(* IEC 61131-3 sources: rsb-lab/vlan50/plc-programs, 6 files *)

(* ---- brewhouse.st ---- *)
PROGRAM plc_prg
VAR
    MashTemp           AT %QW0 : INT;
    MashLevel          AT %QW1 : INT;
    MashPH             AT %QW2 : INT;
    LauterTurbidity    AT %QW3 : INT;
    LauterLevel        AT %QW4 : INT;
    KettleTemp         AT %QW5 : INT;
    KettleLevel        AT %QW6 : INT;
    KettlePressure     AT %QW7 : INT;
    WhirlpoolTemp      AT %QW8 : INT;
    ChillerOutTemp     AT %QW9 : INT;

    MashAgitator       AT %QX0.0 : BOOL;
    MashOutlet         AT %QX0.1 : BOOL;
    LauterToKettle     AT %QX0.2 : BOOL;
    LauterRecirculate  AT %QX0.3 : BOOL;
    KettleSteam        AT %QX0.4 : BOOL;
    KettleToWhirlpool  AT %QX0.5 : BOOL;
    WhirlpoolOutlet    AT %QX0.6 : BOOL;
    ChillerOutlet      AT %QX0.7 : BOOL;

    AlarmTurbidity     AT %QX1.0 : BOOL;  (* coil 8 *)
    AlarmKettleTemp    AT %QX1.1 : BOOL;  (* coil 9 *)
    AlarmKettlePress   AT %QX1.2 : BOOL;  (* coil 10 *)
    AlarmChillerTemp   AT %QX1.3 : BOOL;  (* coil 11 *)
    WhirlpoolReady     AT %QX1.4 : BOOL;  (* coil 12 *)
END_VAR
VAR
    TransferSeen : BOOL;
    WhirlpoolRest : TON;
END_VAR

AlarmTurbidity   := LauterTurbidity > 200;
AlarmKettleTemp  := KettleTemp >= 1000;
AlarmKettlePress := KettlePressure >= 1200;
AlarmChillerTemp := ChillerOutTemp > 200;

IF AlarmTurbidity AND (LauterLevel > 2) THEN
    LauterToKettle := FALSE;
    LauterRecirculate := TRUE;
ELSIF LauterLevel <= 2 THEN
    LauterToKettle := FALSE;
    LauterRecirculate := FALSE;
END_IF;

IF AlarmKettleTemp OR AlarmKettlePress THEN
    KettleSteam := FALSE;
END_IF;

IF KettleToWhirlpool THEN
    TransferSeen := TRUE;
END_IF;

WhirlpoolRest(IN := TransferSeen AND NOT KettleToWhirlpool, PT := T#20m);
WhirlpoolReady := WhirlpoolRest.Q;

IF NOT WhirlpoolReady THEN
    WhirlpoolOutlet := FALSE;
END_IF;

IF AlarmChillerTemp THEN
    ChillerOutlet := FALSE;
END_IF;

IF ChillerOutlet AND (ChillerOutTemp <= 200) THEN
    TransferSeen := FALSE;
END_IF;

END_PROGRAM

CONFIGURATION Config0
    RESOURCE Res0 ON PLC
        TASK task0(INTERVAL := T#100ms, PRIORITY := 0);
        PROGRAM instance0 WITH task0 : plc_prg;
    END_RESOURCE
END_CONFIGURATION

(* ---- conditioning.st ---- *)
PROGRAM plc_prg
VAR
    BBT1Temp       AT %QW0 : INT;
    BBT1Pressure   AT %QW1 : INT;
    BBT1Level      AT %QW2 : INT;
    BBT1Turbidity  AT %QW3 : INT;
    BBT2Temp       AT %QW10 : INT;
    BBT2Pressure   AT %QW11 : INT;
    BBT2Level      AT %QW12 : INT;
    BBT2Turbidity  AT %QW13 : INT;

    BBT1Glycol     AT %QX0.0 : BOOL;
    BBT1CO2Dose    AT %QX0.1 : BOOL;
    BBT1Outlet     AT %QX0.2 : BOOL;
    BBT1Vent       AT %QX0.3 : BOOL;
    BBT2Glycol     AT %QX1.2 : BOOL;
    BBT2CO2Dose    AT %QX1.3 : BOOL;
    BBT2Outlet     AT %QX1.4 : BOOL;
    BBT2Vent       AT %QX1.5 : BOOL;

    AlarmBBT1Temp      AT %QX2.4 : BOOL; (* coil 20 *)
    AlarmBBT2Temp      AT %QX2.5 : BOOL; (* coil 21 *)
    AlarmBBT1Pressure  AT %QX2.6 : BOOL; (* coil 22 *)
    AlarmBBT2Pressure  AT %QX2.7 : BOOL; (* coil 23 *)
    BBT1Ready          AT %QX3.0 : BOOL; (* coil 24 *)
    BBT2Ready          AT %QX3.1 : BOOL; (* coil 25 *)
END_VAR
VAR
    BBT1StableTimer : TON;
    BBT2StableTimer : TON;
END_VAR

AlarmBBT1Temp := BBT1Temp > 20;
AlarmBBT2Temp := BBT2Temp > 20;
AlarmBBT1Pressure := BBT1Pressure > 2000;
AlarmBBT2Pressure := BBT2Pressure > 2000;

IF BBT1Temp > 20 THEN BBT1Glycol := TRUE; ELSIF BBT1Temp <= 0 THEN BBT1Glycol := FALSE; END_IF;
IF BBT2Temp > 20 THEN BBT2Glycol := TRUE; ELSIF BBT2Temp <= 0 THEN BBT2Glycol := FALSE; END_IF;

IF BBT1Pressure > 2000 THEN BBT1CO2Dose := FALSE; END_IF;
IF BBT2Pressure > 2000 THEN BBT2CO2Dose := FALSE; END_IF;

IF BBT1Pressure >= 2500 THEN BBT1Vent := TRUE; ELSIF BBT1Pressure < 2200 THEN BBT1Vent := FALSE; END_IF;
IF BBT2Pressure >= 2500 THEN BBT2Vent := TRUE; ELSIF BBT2Pressure < 2200 THEN BBT2Vent := FALSE; END_IF;

BBT1StableTimer(IN := (BBT1Temp >= 0) AND (BBT1Temp <= 20) AND (BBT1Turbidity <= 20), PT := T#10m);
BBT2StableTimer(IN := (BBT2Temp >= 0) AND (BBT2Temp <= 20) AND (BBT2Turbidity <= 20), PT := T#10m);
BBT1Ready := BBT1StableTimer.Q;
BBT2Ready := BBT2StableTimer.Q;

IF NOT BBT1Ready THEN BBT1Outlet := FALSE; END_IF;
IF NOT BBT2Ready THEN BBT2Outlet := FALSE; END_IF;

IF BBT1Level <= 2 THEN BBT1Outlet := FALSE; END_IF;
IF BBT2Level <= 2 THEN BBT2Outlet := FALSE; END_IF;

END_PROGRAM

CONFIGURATION Config0
    RESOURCE Res0 ON PLC
        TASK task0(INTERVAL := T#100ms, PRIORITY := 0);
        PROGRAM instance0 WITH task0 : plc_prg;
    END_RESOURCE
END_CONFIGURATION

(* ---- fermentation.st ---- *)
PROGRAM plc_prg
VAR
    T1Temp       AT %QW0 : INT;
    T1Pressure   AT %QW1 : INT;
    T1Level      AT %QW2 : INT;
    T1PH         AT %QW3 : INT;
    CO2Header    AT %QW4 : INT;
    CO2Flow      AT %QW5 : INT;

    T2Temp       AT %QW10 : INT;
    T2Pressure   AT %QW11 : INT;
    T2Level      AT %QW12 : INT;
    T2PH         AT %QW13 : INT;
    T3Temp       AT %QW20 : INT;
    T3Pressure   AT %QW21 : INT;
    T3Level      AT %QW22 : INT;
    T3PH         AT %QW23 : INT;
    T4Temp       AT %QW30 : INT;
    T4Pressure   AT %QW31 : INT;
    T4Level      AT %QW32 : INT;
    T4PH         AT %QW33 : INT;

    T1Glycol     AT %QX0.0 : BOOL;
    T1Outlet     AT %QX0.1 : BOOL;
    T1CIP        AT %QX0.2 : BOOL;
    T2Glycol     AT %QX1.2 : BOOL;
    T2Outlet     AT %QX1.3 : BOOL;
    T2CIP        AT %QX1.4 : BOOL;
    T3Glycol     AT %QX2.4 : BOOL;
    T3Outlet     AT %QX2.5 : BOOL;
    T3CIP        AT %QX2.6 : BOOL;
    T4Glycol     AT %QX3.6 : BOOL;
    T4Outlet     AT %QX3.7 : BOOL;
    T4CIP        AT %QX4.0 : BOOL;
    CO2Vent      AT %QX5.0 : BOOL;
    CO2Recovery  AT %QX5.1 : BOOL;

    AlarmHighPressure AT %QX6.2 : BOOL; (* coil 50 *)
    AlarmEmergency    AT %QX6.3 : BOOL; (* coil 51 *)
    T1Complete        AT %QX6.4 : BOOL; (* coil 52 *)
    T2Complete        AT %QX6.5 : BOOL; (* coil 53 *)
    T3Complete        AT %QX6.6 : BOOL; (* coil 54 *)
    T4Complete        AT %QX6.7 : BOOL; (* coil 55 *)
END_VAR
VAR
    T1FermentTimer : TON;
    T2FermentTimer : TON;
    T3FermentTimer : TON;
    T4FermentTimer : TON;
END_VAR

IF T1Temp > 205 THEN T1Glycol := TRUE; ELSIF T1Temp < 195 THEN T1Glycol := FALSE; END_IF;
IF T2Temp > 205 THEN T2Glycol := TRUE; ELSIF T2Temp < 195 THEN T2Glycol := FALSE; END_IF;
IF T3Temp > 205 THEN T3Glycol := TRUE; ELSIF T3Temp < 195 THEN T3Glycol := FALSE; END_IF;
IF T4Temp > 205 THEN T4Glycol := TRUE; ELSIF T4Temp < 195 THEN T4Glycol := FALSE; END_IF;

AlarmHighPressure := (T1Pressure > 1500) OR (T2Pressure > 1500) OR
                     (T3Pressure > 1500) OR (T4Pressure > 1500);
AlarmEmergency := (T1Pressure > 2000) OR (T2Pressure > 2000) OR
                  (T3Pressure > 2000) OR (T4Pressure > 2000);

IF AlarmHighPressure THEN
    CO2Vent := TRUE;
ELSIF (T1Pressure < 1350) AND (T2Pressure < 1350) AND
      (T3Pressure < 1350) AND (T4Pressure < 1350) THEN
    CO2Vent := FALSE;
END_IF;

IF AlarmEmergency THEN
    T1CIP := FALSE;
    T2CIP := FALSE;
    T3CIP := FALSE;
    T4CIP := FALSE;
END_IF;

IF CO2Header > 1200 AND NOT CO2Vent THEN
    CO2Recovery := TRUE;
ELSIF CO2Header < 1100 OR CO2Vent THEN
    CO2Recovery := FALSE;
END_IF;

T1FermentTimer(IN := T1PH <= 420, PT := T#10m);
T2FermentTimer(IN := T2PH <= 420, PT := T#10m);
T3FermentTimer(IN := T3PH <= 420, PT := T#10m);
T4FermentTimer(IN := T4PH <= 420, PT := T#10m);
T1Complete := T1FermentTimer.Q;
T2Complete := T2FermentTimer.Q;
T3Complete := T3FermentTimer.Q;
T4Complete := T4FermentTimer.Q;

IF (NOT T1Complete) OR T1CIP THEN T1Outlet := FALSE; END_IF;
IF (NOT T2Complete) OR T2CIP THEN T2Outlet := FALSE; END_IF;
IF (NOT T3Complete) OR T3CIP THEN T3Outlet := FALSE; END_IF;
IF (NOT T4Complete) OR T4CIP THEN T4Outlet := FALSE; END_IF;

END_PROGRAM

CONFIGURATION Config0
    RESOURCE Res0 ON PLC
        TASK task0(INTERVAL := T#100ms, PRIORITY := 0);
        PROGRAM instance0 WITH task0 : plc_prg;
    END_RESOURCE
END_CONFIGURATION

(* ---- packaging.st ---- *)
PROGRAM plc_prg
VAR
    FilterDP       AT %QW0 : INT;
    FlowRate       AT %QW1 : INT;
    SourceLevel    AT %QW2 : INT;
    BottleCount    AT %QW3 : INT;
    CapTorque      AT %QW4 : INT;
    CaseCount      AT %QW5 : INT;

    FillerRun      AT %QX0.0 : BOOL;
    CIPActive      AT %QX0.1 : BOOL;
    CapperRun      AT %QX0.2 : BOOL;
    ConveyorZ1     AT %QX0.3 : BOOL;
    ConveyorZ2     AT %QX0.4 : BOOL;
    ConveyorZ3     AT %QX0.5 : BOOL;
    LineEStop      AT %QX0.6 : BOOL;
    RejectGate     AT %QX0.7 : BOOL;

    AlarmLowFlow   AT %QX1.0 : BOOL; (* coil 8 *)
    AlarmCapTorque AT %QX1.1 : BOOL; (* coil 9 *)
    AlarmFilterDP  AT %QX1.2 : BOOL; (* coil 10 *)
    AlarmLowLevel  AT %QX1.3 : BOOL; (* coil 11 *)
END_VAR
VAR
    FillerStartup : TON;
END_VAR

FillerStartup(IN := FillerRun AND NOT CIPActive AND NOT LineEStop, PT := T#10s);
AlarmLowFlow := FillerStartup.Q AND (FlowRate < 5);
AlarmCapTorque := FillerRun AND CapperRun AND ((CapTorque < 20) OR (CapTorque > 40));
AlarmFilterDP := FilterDP >= 400;
AlarmLowLevel := SourceLevel <= 5;
RejectGate := AlarmCapTorque;

IF CIPActive THEN
    FillerRun := FALSE;
    CapperRun := FALSE;
    ConveyorZ1 := FALSE;
    ConveyorZ2 := FALSE;
    ConveyorZ3 := FALSE;
END_IF;

IF AlarmLowFlow OR AlarmLowLevel THEN
    FillerRun := FALSE;
END_IF;

IF AlarmFilterDP THEN
    LineEStop := TRUE;
END_IF;

IF LineEStop THEN
    FillerRun := FALSE;
    CapperRun := FALSE;
    ConveyorZ1 := FALSE;
    ConveyorZ2 := FALSE;
    ConveyorZ3 := FALSE;
END_IF;

END_PROGRAM

CONFIGURATION Config0
    RESOURCE Res0 ON PLC
        TASK task0(INTERVAL := T#100ms, PRIORITY := 0);
        PROGRAM instance0 WITH task0 : plc_prg;
    END_RESOURCE
END_CONFIGURATION

(* ---- rawmat.st ---- *)
PROGRAM plc_prg
VAR
    Silo1_kg       AT %QW0 : INT;
    Silo2_kg       AT %QW1 : INT;
    MillRPM        AT %QW2 : INT;
    AugerCurrent   AT %QW3 : INT;
    HLT_Temp       AT %QW4 : INT;
    HLT_Level      AT %QW5 : INT;
    HLT_Flow       AT %QW6 : INT;
    CLT_Temp       AT %QW7 : INT;
    CLT_Level      AT %QW8 : INT;

    MillMotor      AT %QX0.0 : BOOL;
    AugerMotor     AT %QX0.1 : BOOL;
    HLT_Heater     AT %QX0.2 : BOOL;
    HLT_Valve      AT %QX0.3 : BOOL;
    CLT_Valve      AT %QX0.4 : BOOL;

    AlarmSiloLow   AT %QX1.0 : BOOL;  (* coil 8 *)
    AlarmAugerJam  AT %QX1.1 : BOOL;  (* coil 9 *)
    AlarmHLTHigh   AT %QX1.2 : BOOL;  (* coil 10 *)
    AlarmTankLow   AT %QX1.3 : BOOL;  (* coil 11 *)
END_VAR

AlarmSiloLow  := (Silo1_kg < 500) AND (Silo2_kg < 500);
AlarmAugerJam := AugerCurrent >= 100;   (* 10.0 A *)
AlarmHLTHigh  := HLT_Temp >= 780;       (* 78.0 C *)
AlarmTankLow  := (HLT_Level <= 5) OR (CLT_Level <= 5);

IF AlarmSiloLow OR AlarmAugerJam THEN
    MillMotor := FALSE;
    AugerMotor := FALSE;
END_IF;

IF AlarmHLTHigh THEN
    HLT_Heater := FALSE;
END_IF;

IF HLT_Level <= 5 THEN
    HLT_Valve := FALSE;
END_IF;

IF CLT_Level <= 5 THEN
    CLT_Valve := FALSE;
END_IF;

END_PROGRAM

CONFIGURATION Config0
    RESOURCE Res0 ON PLC
        TASK task0(INTERVAL := T#100ms, PRIORITY := 0);
        PROGRAM instance0 WITH task0 : plc_prg;
    END_RESOURCE
END_CONFIGURATION

(* ---- utilities.st ---- *)
PROGRAM plc_prg
VAR
    AirPressure       AT %QW0 : INT;
    AirDewPoint       AT %QW1 : INT;
    CO2Pressure       AT %QW2 : INT;
    CO2Level          AT %QW3 : INT;
    Conductivity      AT %QW4 : INT;
    UVLampOK          AT %QW5 : INT;

    BoilerDrumPress   AT %QW700 : INT;
    SteamHeaderPress  AT %QW701 : INT;
    FlueTemp          AT %QW702 : INT;
    FeedWaterLevel    AT %QW703 : INT;
    BurnerStatus      AT %QW704 : INT;
    ReliefStatus      AT %QW705 : INT;

    BurnerEnable      AT %QX0.0 : BOOL;
    FeedPump          AT %QX0.1 : BOOL;
    AirHeaderValve    AT %QX0.2 : BOOL;
    CO2Regulator      AT %QX0.3 : BOOL;
    WaterOutlet       AT %QX0.4 : BOOL;

    AlarmBoilerTrip   AT %QX1.0 : BOOL; (* coil 8 *)
    AlarmAirLow       AT %QX1.1 : BOOL; (* coil 9 *)
    AlarmCO2Low       AT %QX1.2 : BOOL; (* coil 10 *)
    AlarmUVFault      AT %QX1.3 : BOOL; (* coil 11 *)
    AlarmSteamLow     AT %QX1.4 : BOOL; (* coil 12 *)
    AlarmWaterQuality AT %QX1.5 : BOOL; (* coil 13 *)
END_VAR

AlarmBoilerTrip := (BoilerDrumPress > 100) OR (FeedWaterLevel < 10);
AlarmSteamLow := SteamHeaderPress < 40;
AlarmAirLow := AirPressure < 50;
AlarmCO2Low := CO2Level < 20;
AlarmUVFault := UVLampOK = 0;
AlarmWaterQuality := Conductivity > 100;

(* Boiler burner demand control.
   Drum pressure register is bar x 10, so 70 = 7.0 bar setpoint.
   Hysteresis band 6.6-7.0 bar lets the burner cycle and hold steam
   pressure instead of staying off from cold start. *)
IF BoilerDrumPress < 66 THEN
    BurnerEnable := TRUE;
ELSIF BoilerDrumPress >= 70 THEN
    BurnerEnable := FALSE;
END_IF;

(* Safety trip always overrides burner demand. *)
IF AlarmBoilerTrip THEN
    BurnerEnable := FALSE;
END_IF;

(* Feed-water level control with hysteresis, kept well above the
   10% low-level trip so the burner interlock stays satisfied. *)
IF FeedWaterLevel < 40 THEN
    FeedPump := TRUE;
ELSIF FeedWaterLevel >= 70 THEN
    FeedPump := FALSE;
END_IF;

IF AlarmCO2Low THEN
    CO2Regulator := FALSE;
END_IF;

IF AlarmUVFault OR AlarmWaterQuality THEN
    WaterOutlet := FALSE;
END_IF;

END_PROGRAM

CONFIGURATION Config0
    RESOURCE Res0 ON PLC
        TASK task0(INTERVAL := T#100ms, PRIORITY := 0);
        PROGRAM instance0 WITH task0 : plc_prg;
    END_RESOURCE
END_CONFIGURATION
